// CFC twin of T_SafeMuting_Tests: the same tests drawn as CFC diagrams, the way a TwinSAFE project is authored.
    FUNCTION_BLOCK T_SafeMuting_Tests_CFC EXTENDS T_SafeCfcTestSuite
    VAR
    // Test_OssdBlockedWithoutMutingGivesSafe
    group_1 : T_SafeGroup;
    fb_1 : T_SafeMuting(group := group_1);
    // Test_SequentialMutingKeepsOutputOn
    group_2 : T_SafeGroup;
    fb_2 : T_SafeMuting(group := group_2) := (Parameters := (SequentialInputs := TRUE));
    // Test_SequenceViolationGivesError
    group_3 : T_SafeGroup;
    fb_3 : T_SafeMuting(group := group_3) := (Parameters := (SequentialInputs := TRUE));
    // Test_TwoSensorParallelSequence
    group_4 : T_SafeGroup;
    fb_4 : T_SafeMuting(group := group_4);
END_VAR

Test_OssdBlockedWithoutMutingGivesSafe();
Test_SequentialMutingKeepsOutputOn();
Test_SequenceViolationGivesError();
Test_TwoSensorParallelSequence();

METHOD PRIVATE Test_OssdBlockedWithoutMutingGivesSafe
// note: this text did not pass the execution check against the stored diagram
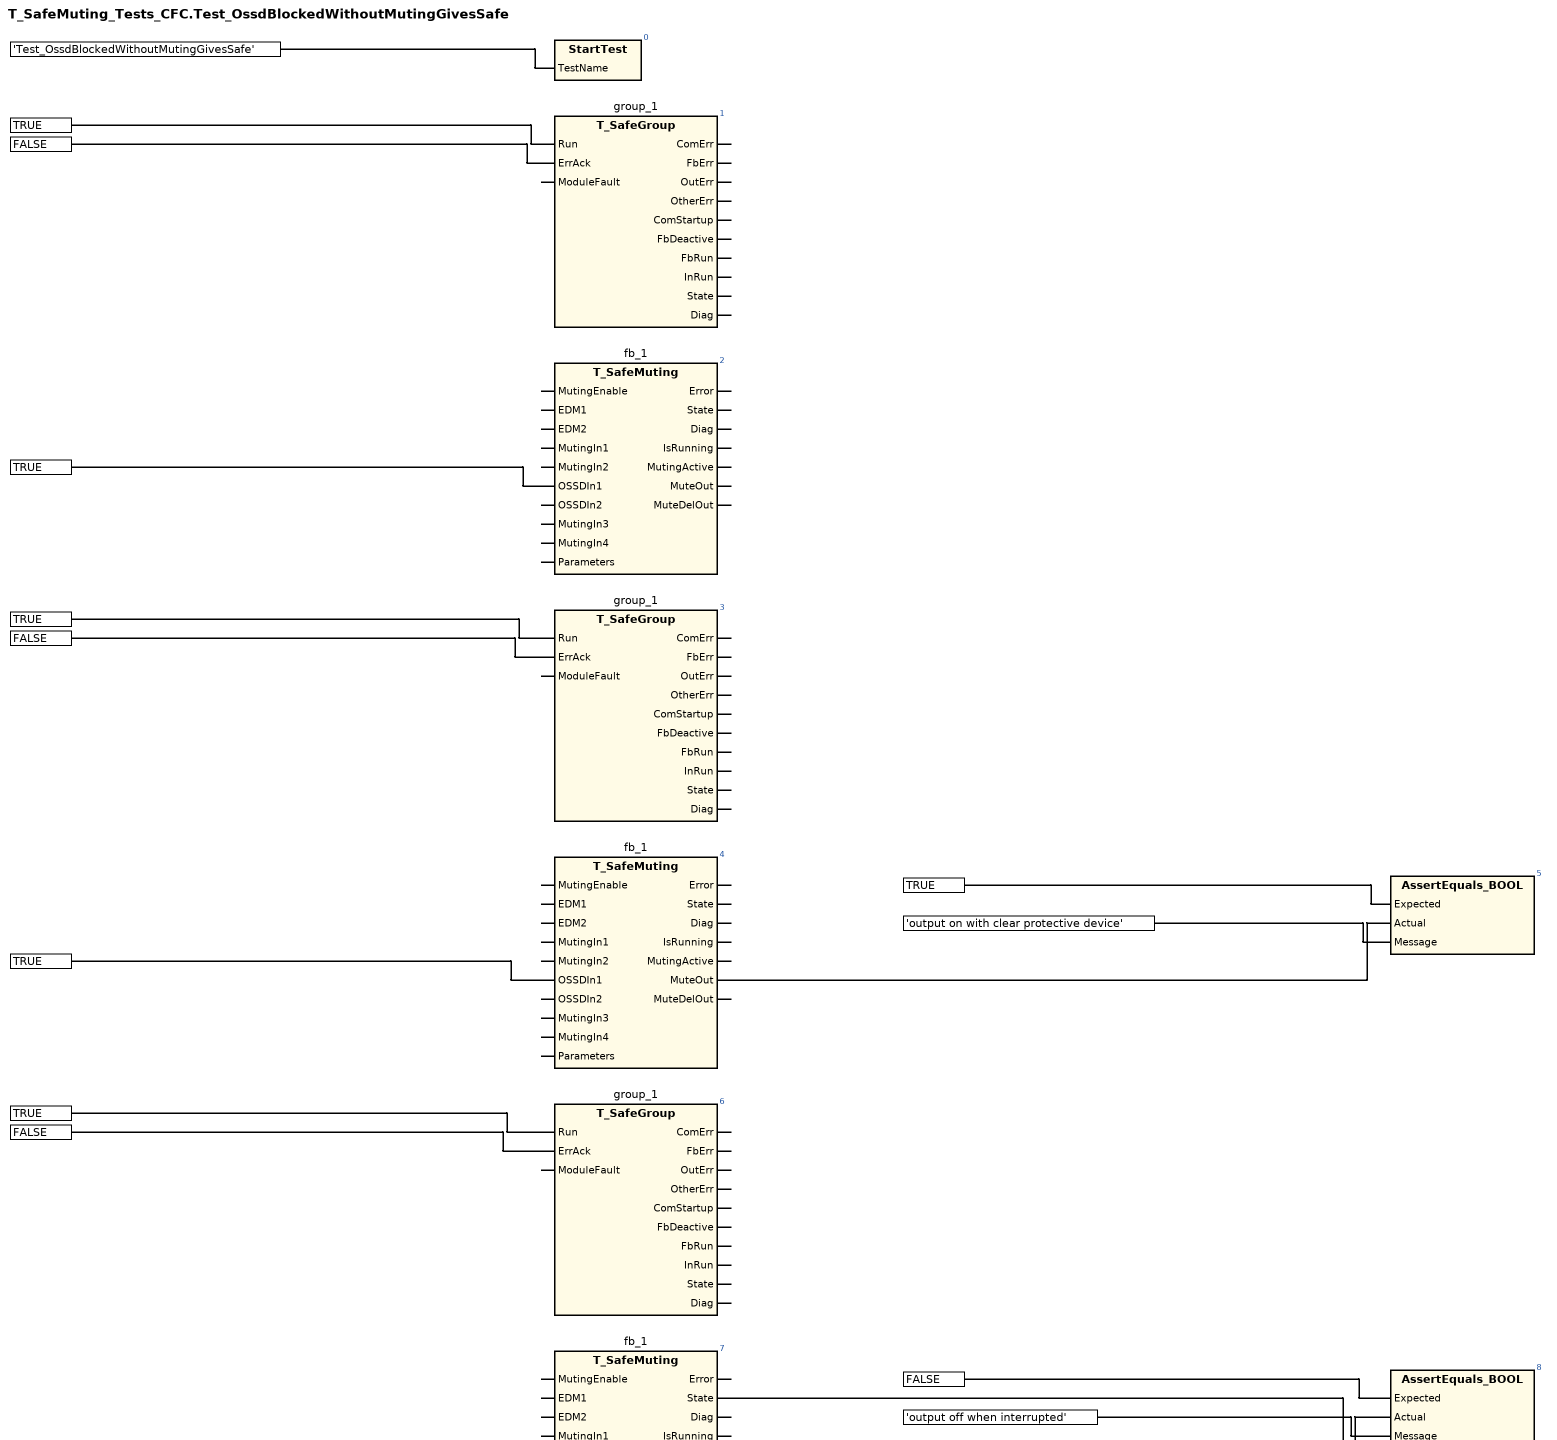
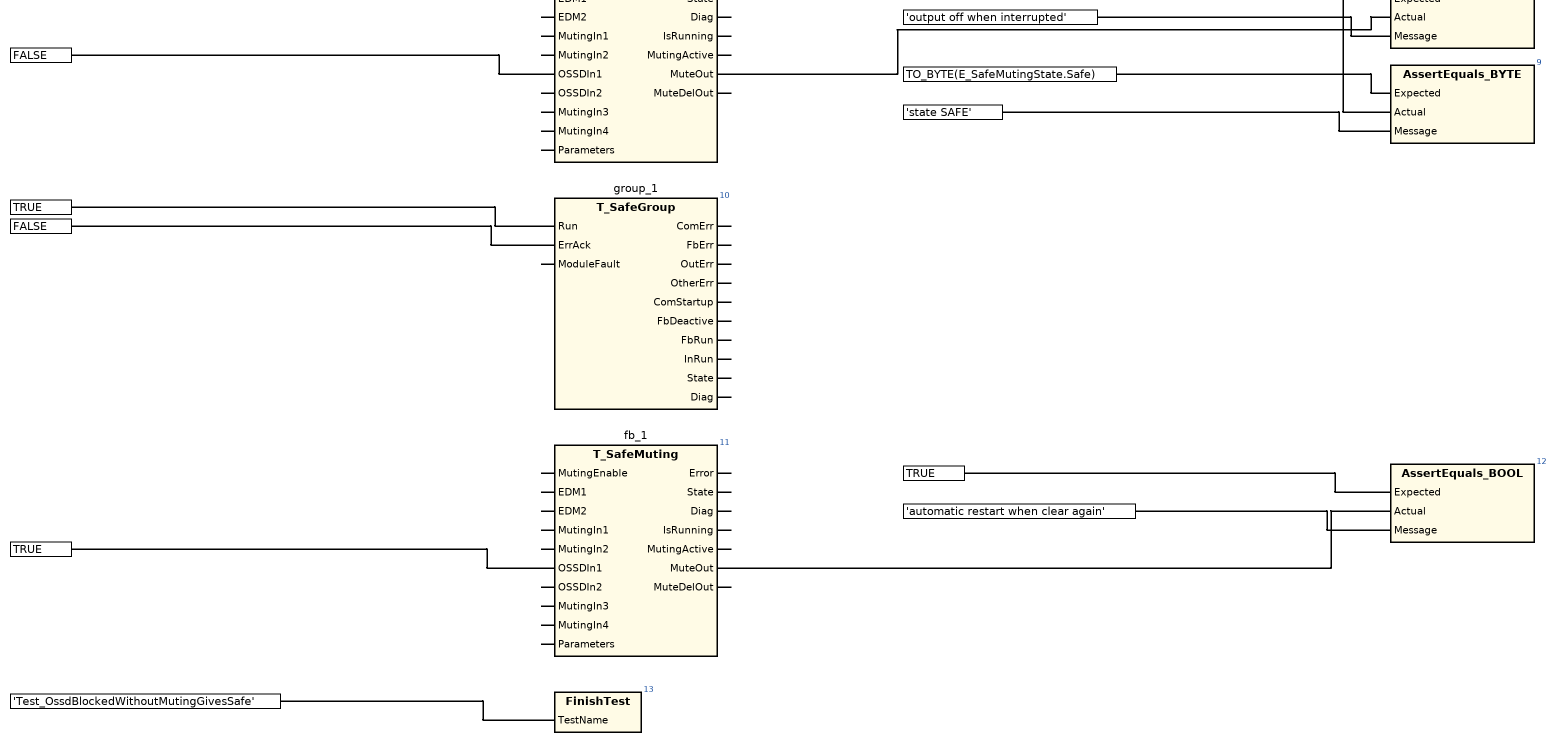
StartTest(TestName := 'Test_OssdBlockedWithoutMutingGivesSafe');
group_1(Run := TRUE, ErrAck := FALSE); // T_SafeGroup
fb_1(OSSDIn1 := TRUE); // T_SafeMuting
group_1(Run := TRUE, ErrAck := FALSE); // T_SafeGroup
fb_1(OSSDIn1 := TRUE); // T_SafeMuting
AssertEquals_BOOL(Expected := TRUE, Actual := fb_1.MuteOut, Message := 'output on with clear protective device');
group_1(Run := TRUE, ErrAck := FALSE); // T_SafeGroup
fb_1(OSSDIn1 := FALSE); // T_SafeMuting
AssertEquals_BOOL(Expected := FALSE, Actual := fb_1.MuteOut, Message := 'output off when interrupted');
AssertEquals_BYTE(Expected := TO_BYTE(E_SafeMutingState.Safe), Actual := fb_1.State, Message := 'state SAFE');
group_1(Run := TRUE, ErrAck := FALSE); // T_SafeGroup
fb_1(OSSDIn1 := TRUE); // T_SafeMuting
AssertEquals_BOOL(Expected := TRUE, Actual := fb_1.MuteOut, Message := 'automatic restart when clear again');
FinishTest(TestName := 'Test_OssdBlockedWithoutMutingGivesSafe');
END_METHOD

METHOD PRIVATE Test_SequentialMutingKeepsOutputOn
// note: this text did not pass the execution check against the stored diagram
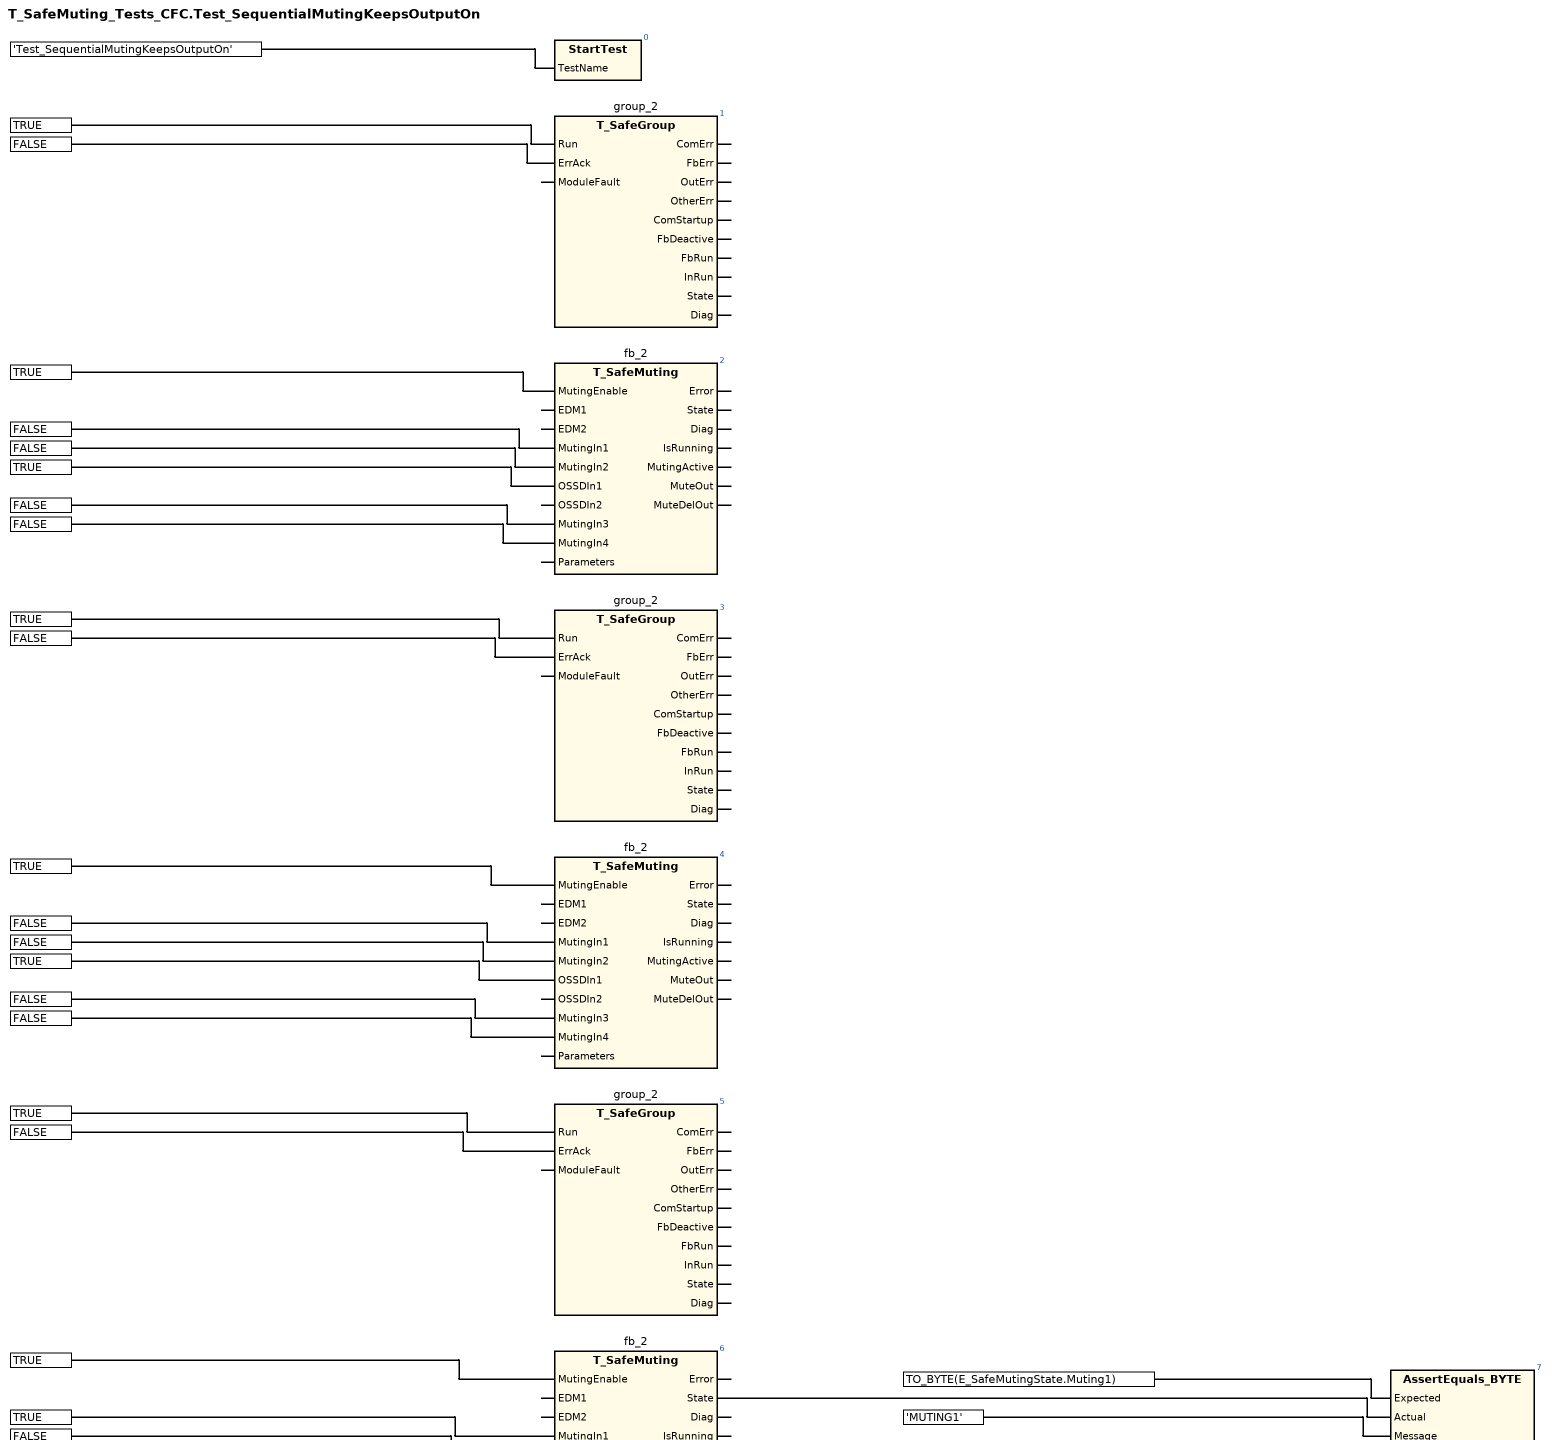
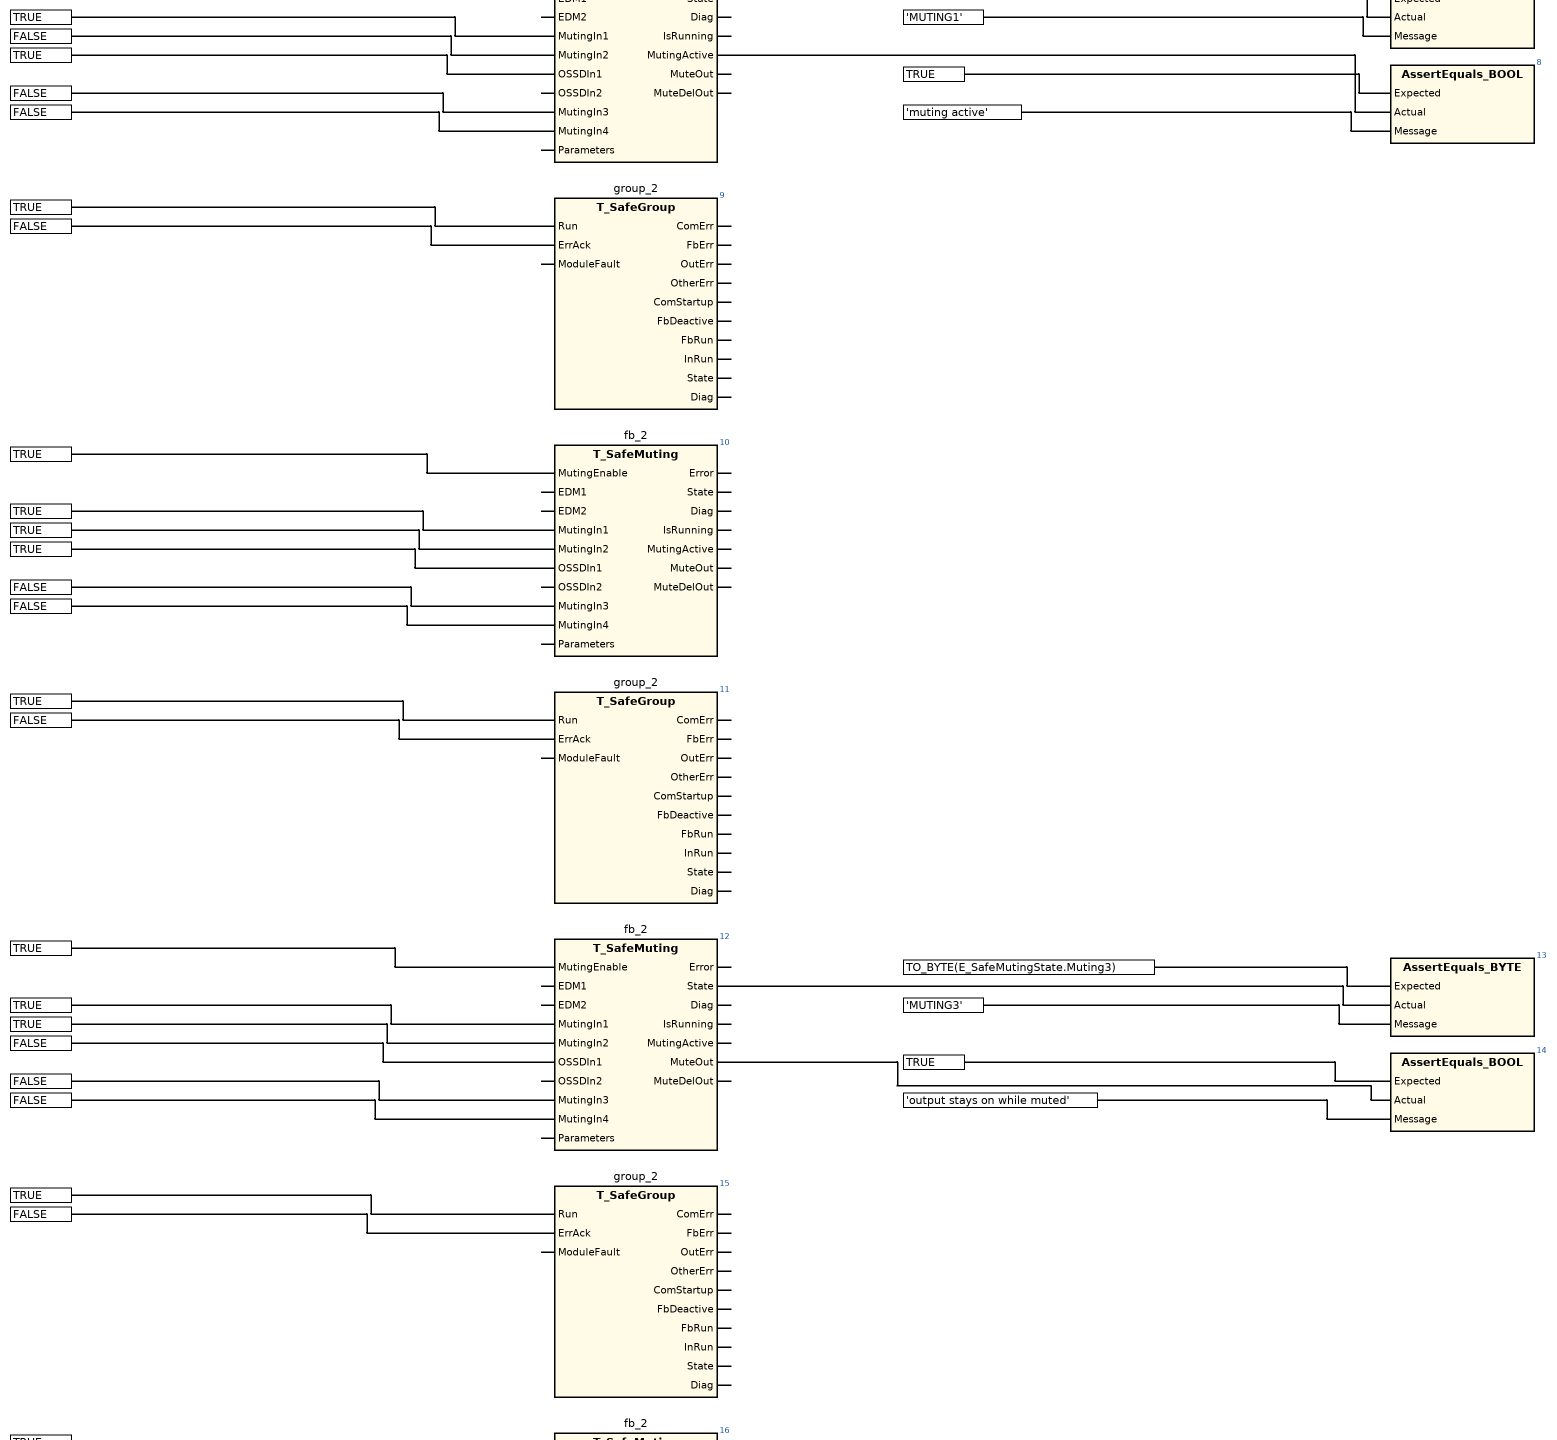
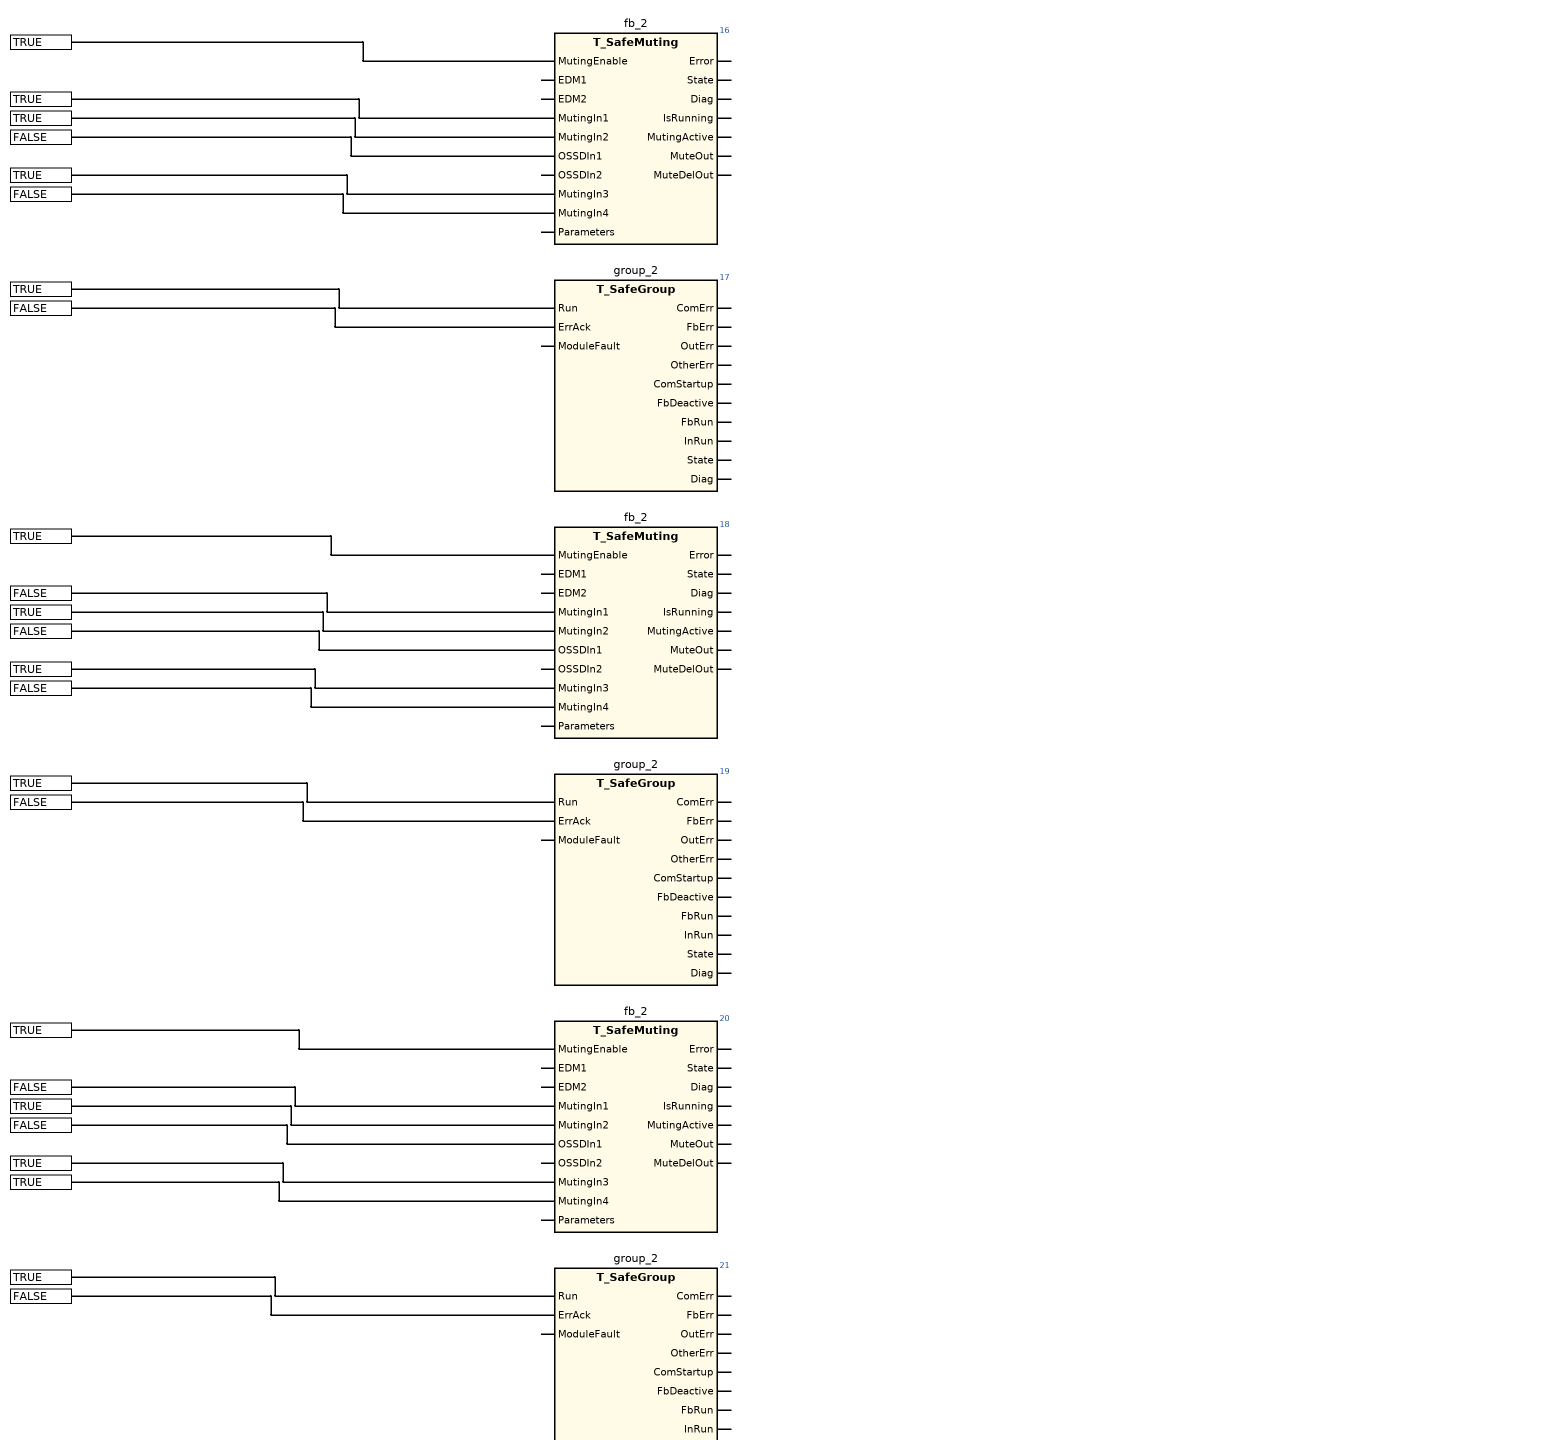
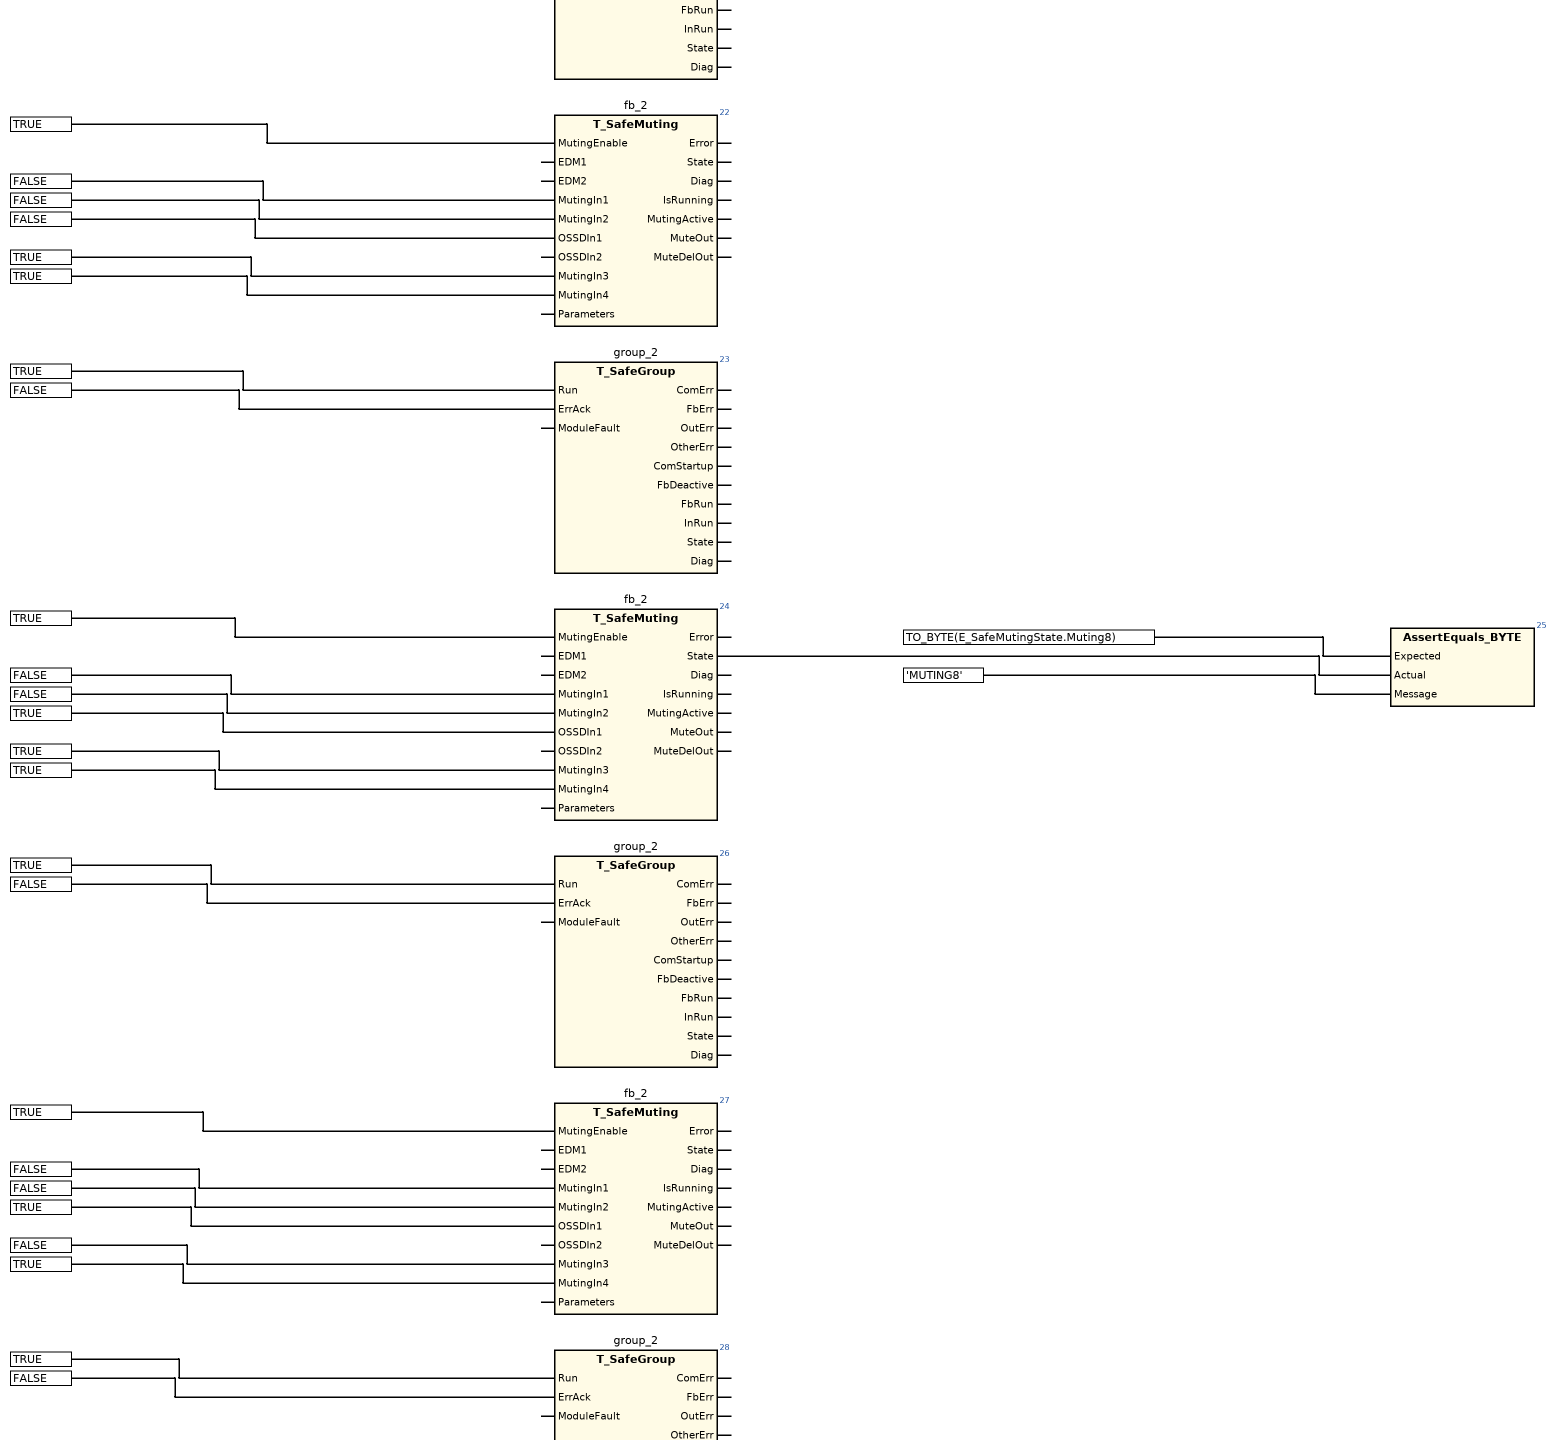
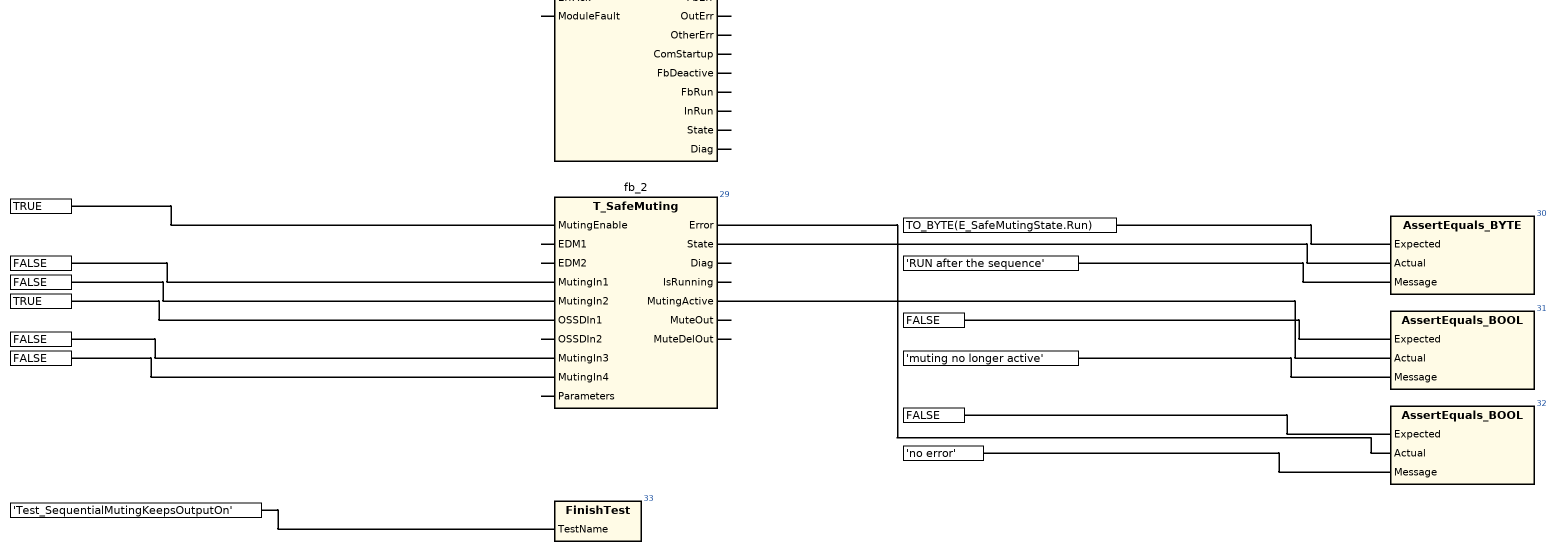
StartTest(TestName := 'Test_SequentialMutingKeepsOutputOn');
group_2(Run := TRUE, ErrAck := FALSE); // T_SafeGroup
fb_2(
    MutingEnable := TRUE,
    MutingIn1 := FALSE,
    MutingIn2 := FALSE,
    OSSDIn1 := TRUE,
    MutingIn3 := FALSE,
    MutingIn4 := FALSE); // T_SafeMuting
group_2(Run := TRUE, ErrAck := FALSE); // T_SafeGroup
fb_2(
    MutingEnable := TRUE,
    MutingIn1 := FALSE,
    MutingIn2 := FALSE,
    OSSDIn1 := TRUE,
    MutingIn3 := FALSE,
    MutingIn4 := FALSE); // T_SafeMuting
group_2(Run := TRUE, ErrAck := FALSE); // T_SafeGroup
fb_2(
    MutingEnable := TRUE,
    MutingIn1 := TRUE,
    MutingIn2 := FALSE,
    OSSDIn1 := TRUE,
    MutingIn3 := FALSE,
    MutingIn4 := FALSE); // T_SafeMuting
AssertEquals_BYTE(Expected := TO_BYTE(E_SafeMutingState.Muting1), Actual := fb_2.State, Message := 'MUTING1');
AssertEquals_BOOL(Expected := TRUE, Actual := fb_2.MutingActive, Message := 'muting active');
group_2(Run := TRUE, ErrAck := FALSE); // T_SafeGroup
fb_2(
    MutingEnable := TRUE,
    MutingIn1 := TRUE,
    MutingIn2 := TRUE,
    OSSDIn1 := TRUE,
    MutingIn3 := FALSE,
    MutingIn4 := FALSE); // T_SafeMuting
group_2(Run := TRUE, ErrAck := FALSE); // T_SafeGroup
fb_2(
    MutingEnable := TRUE,
    MutingIn1 := TRUE,
    MutingIn2 := TRUE,
    OSSDIn1 := FALSE,
    MutingIn3 := FALSE,
    MutingIn4 := FALSE); // T_SafeMuting
AssertEquals_BYTE(Expected := TO_BYTE(E_SafeMutingState.Muting3), Actual := fb_2.State, Message := 'MUTING3');
AssertEquals_BOOL(Expected := TRUE, Actual := fb_2.MuteOut, Message := 'output stays on while muted');
group_2(Run := TRUE, ErrAck := FALSE); // T_SafeGroup
fb_2(
    MutingEnable := TRUE,
    MutingIn1 := TRUE,
    MutingIn2 := TRUE,
    OSSDIn1 := FALSE,
    MutingIn3 := TRUE,
    MutingIn4 := FALSE); // T_SafeMuting
group_2(Run := TRUE, ErrAck := FALSE); // T_SafeGroup
fb_2(
    MutingEnable := TRUE,
    MutingIn1 := FALSE,
    MutingIn2 := TRUE,
    OSSDIn1 := FALSE,
    MutingIn3 := TRUE,
    MutingIn4 := FALSE); // T_SafeMuting
group_2(Run := TRUE, ErrAck := FALSE); // T_SafeGroup
fb_2(
    MutingEnable := TRUE,
    MutingIn1 := FALSE,
    MutingIn2 := TRUE,
    OSSDIn1 := FALSE,
    MutingIn3 := TRUE,
    MutingIn4 := TRUE); // T_SafeMuting
group_2(Run := TRUE, ErrAck := FALSE); // T_SafeGroup
fb_2(
    MutingEnable := TRUE,
    MutingIn1 := FALSE,
    MutingIn2 := FALSE,
    OSSDIn1 := FALSE,
    MutingIn3 := TRUE,
    MutingIn4 := TRUE); // T_SafeMuting
group_2(Run := TRUE, ErrAck := FALSE); // T_SafeGroup
fb_2(
    MutingEnable := TRUE,
    MutingIn1 := FALSE,
    MutingIn2 := FALSE,
    OSSDIn1 := TRUE,
    MutingIn3 := TRUE,
    MutingIn4 := TRUE); // T_SafeMuting
AssertEquals_BYTE(Expected := TO_BYTE(E_SafeMutingState.Muting8), Actual := fb_2.State, Message := 'MUTING8');
group_2(Run := TRUE, ErrAck := FALSE); // T_SafeGroup
fb_2(
    MutingEnable := TRUE,
    MutingIn1 := FALSE,
    MutingIn2 := FALSE,
    OSSDIn1 := TRUE,
    MutingIn3 := FALSE,
    MutingIn4 := TRUE); // T_SafeMuting
group_2(Run := TRUE, ErrAck := FALSE); // T_SafeGroup
fb_2(
    MutingEnable := TRUE,
    MutingIn1 := FALSE,
    MutingIn2 := FALSE,
    OSSDIn1 := TRUE,
    MutingIn3 := FALSE,
    MutingIn4 := FALSE); // T_SafeMuting
AssertEquals_BYTE(Expected := TO_BYTE(E_SafeMutingState.Run), Actual := fb_2.State, Message := 'RUN after the sequence');
AssertEquals_BOOL(Expected := FALSE, Actual := fb_2.MutingActive, Message := 'muting no longer active');
AssertEquals_BOOL(Expected := FALSE, Actual := fb_2.Error, Message := 'no error');
FinishTest(TestName := 'Test_SequentialMutingKeepsOutputOn');
END_METHOD

METHOD PRIVATE Test_SequenceViolationGivesError
// note: this text did not pass the execution check against the stored diagram
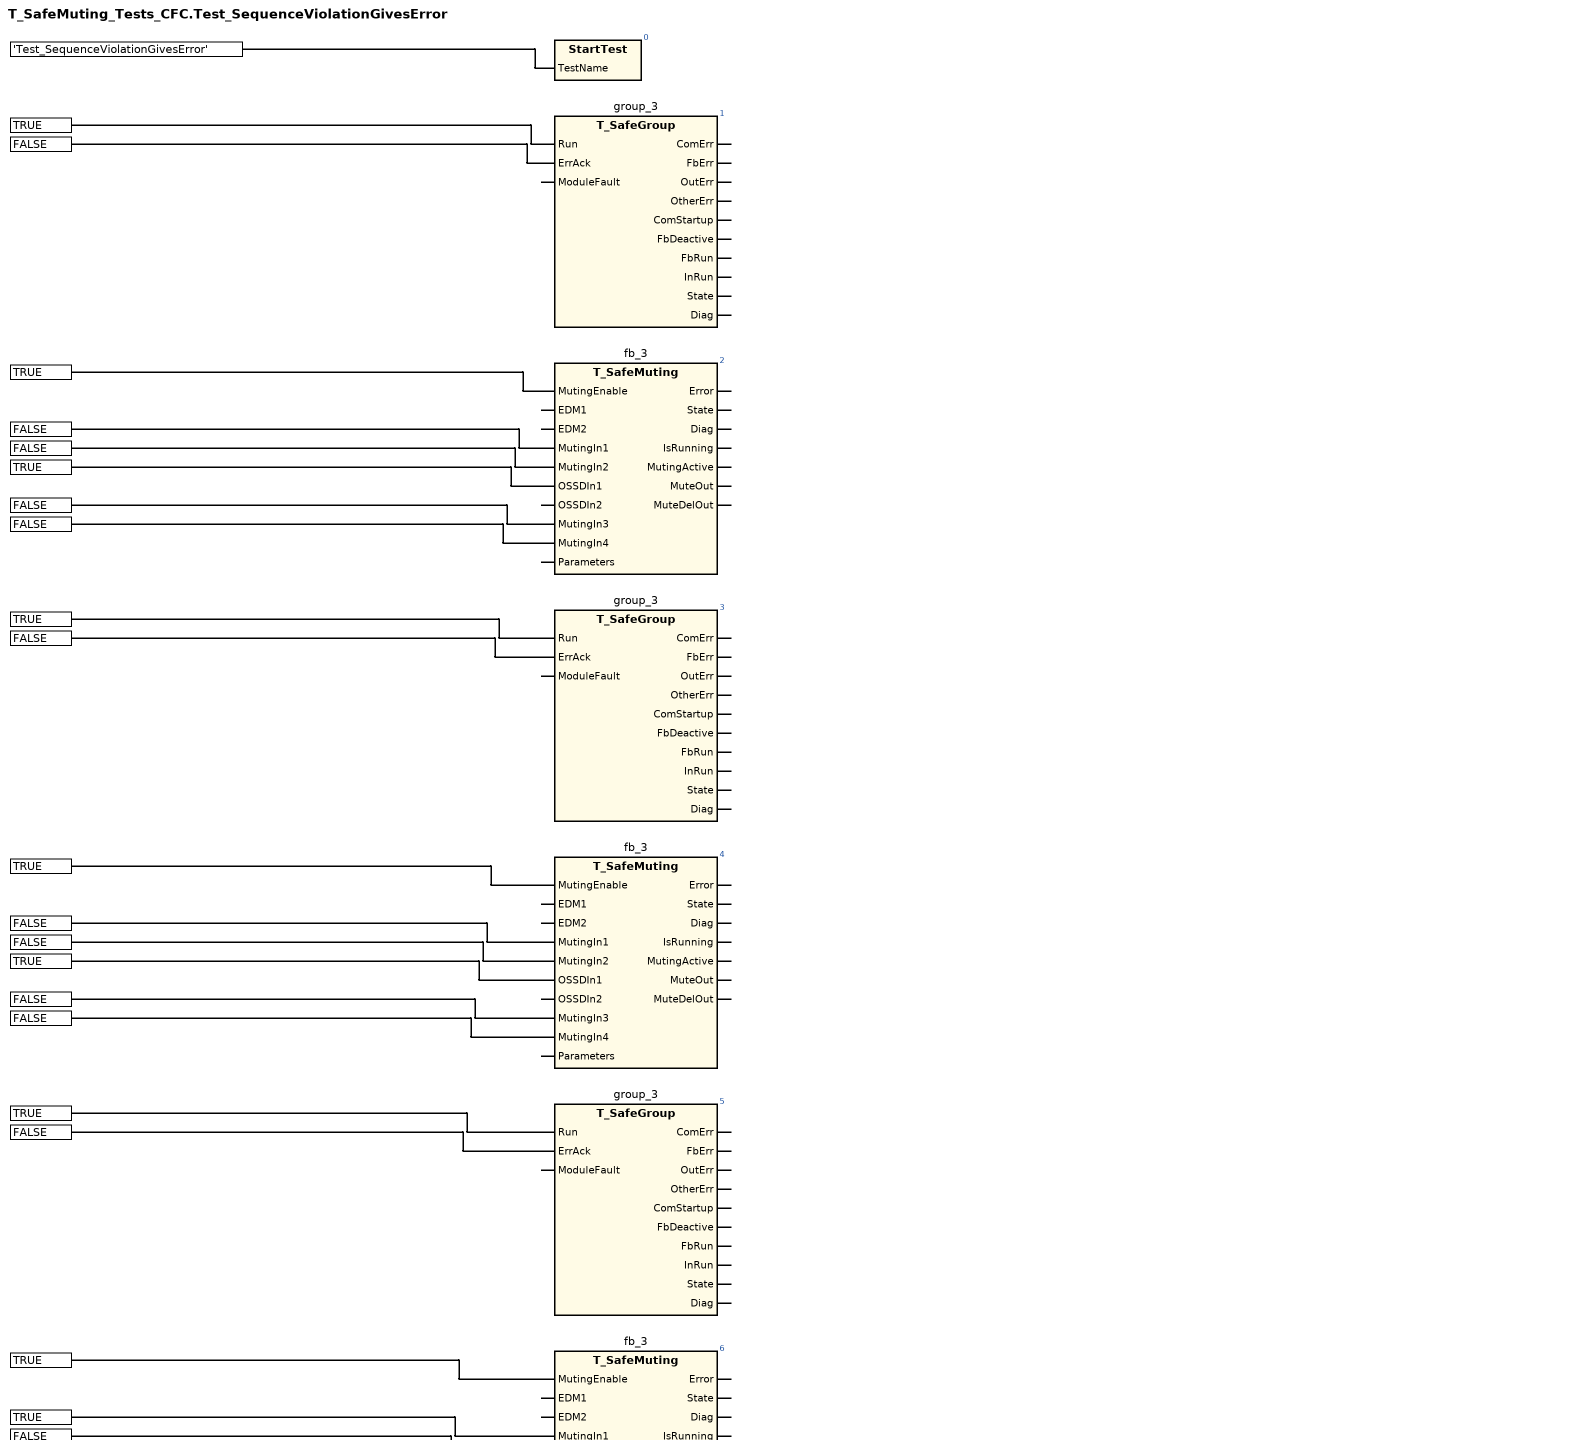
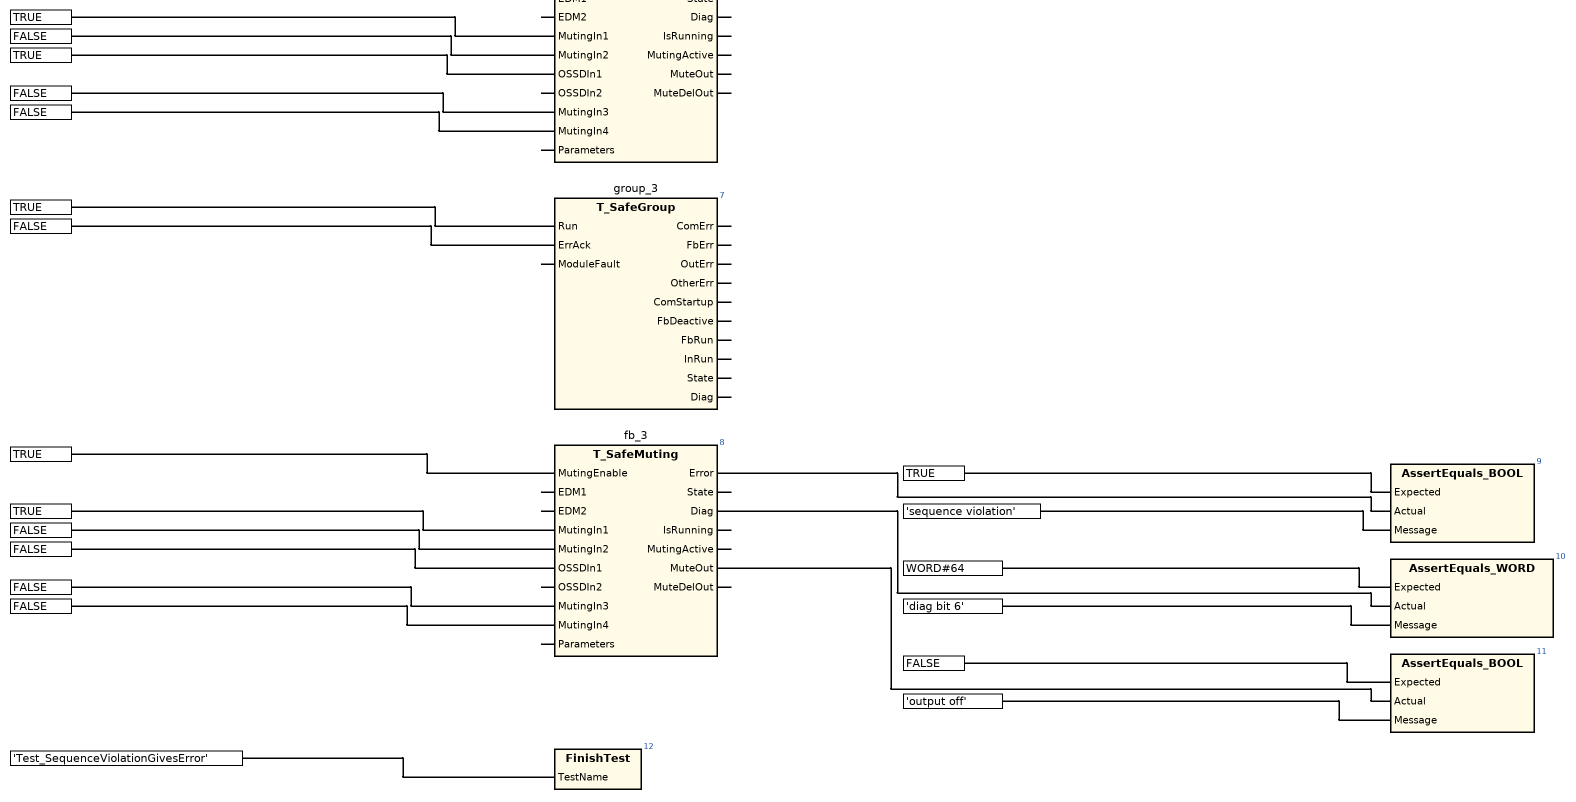
StartTest(TestName := 'Test_SequenceViolationGivesError');
group_3(Run := TRUE, ErrAck := FALSE); // T_SafeGroup
fb_3(
    MutingEnable := TRUE,
    MutingIn1 := FALSE,
    MutingIn2 := FALSE,
    OSSDIn1 := TRUE,
    MutingIn3 := FALSE,
    MutingIn4 := FALSE); // T_SafeMuting
group_3(Run := TRUE, ErrAck := FALSE); // T_SafeGroup
fb_3(
    MutingEnable := TRUE,
    MutingIn1 := FALSE,
    MutingIn2 := FALSE,
    OSSDIn1 := TRUE,
    MutingIn3 := FALSE,
    MutingIn4 := FALSE); // T_SafeMuting
group_3(Run := TRUE, ErrAck := FALSE); // T_SafeGroup
fb_3(
    MutingEnable := TRUE,
    MutingIn1 := TRUE,
    MutingIn2 := FALSE,
    OSSDIn1 := TRUE,
    MutingIn3 := FALSE,
    MutingIn4 := FALSE); // T_SafeMuting
group_3(Run := TRUE, ErrAck := FALSE); // T_SafeGroup
fb_3(
    MutingEnable := TRUE,
    MutingIn1 := TRUE,
    MutingIn2 := FALSE,
    OSSDIn1 := FALSE,
    MutingIn3 := FALSE,
    MutingIn4 := FALSE); // T_SafeMuting
AssertEquals_BOOL(Expected := TRUE, Actual := fb_3.Error, Message := 'sequence violation');
AssertEquals_WORD(Expected := WORD#64, Actual := fb_3.Diag, Message := 'diag bit 6');
AssertEquals_BOOL(Expected := FALSE, Actual := fb_3.MuteOut, Message := 'output off');
FinishTest(TestName := 'Test_SequenceViolationGivesError');
END_METHOD

METHOD PRIVATE Test_TwoSensorParallelSequence
// note: this text did not pass the execution check against the stored diagram
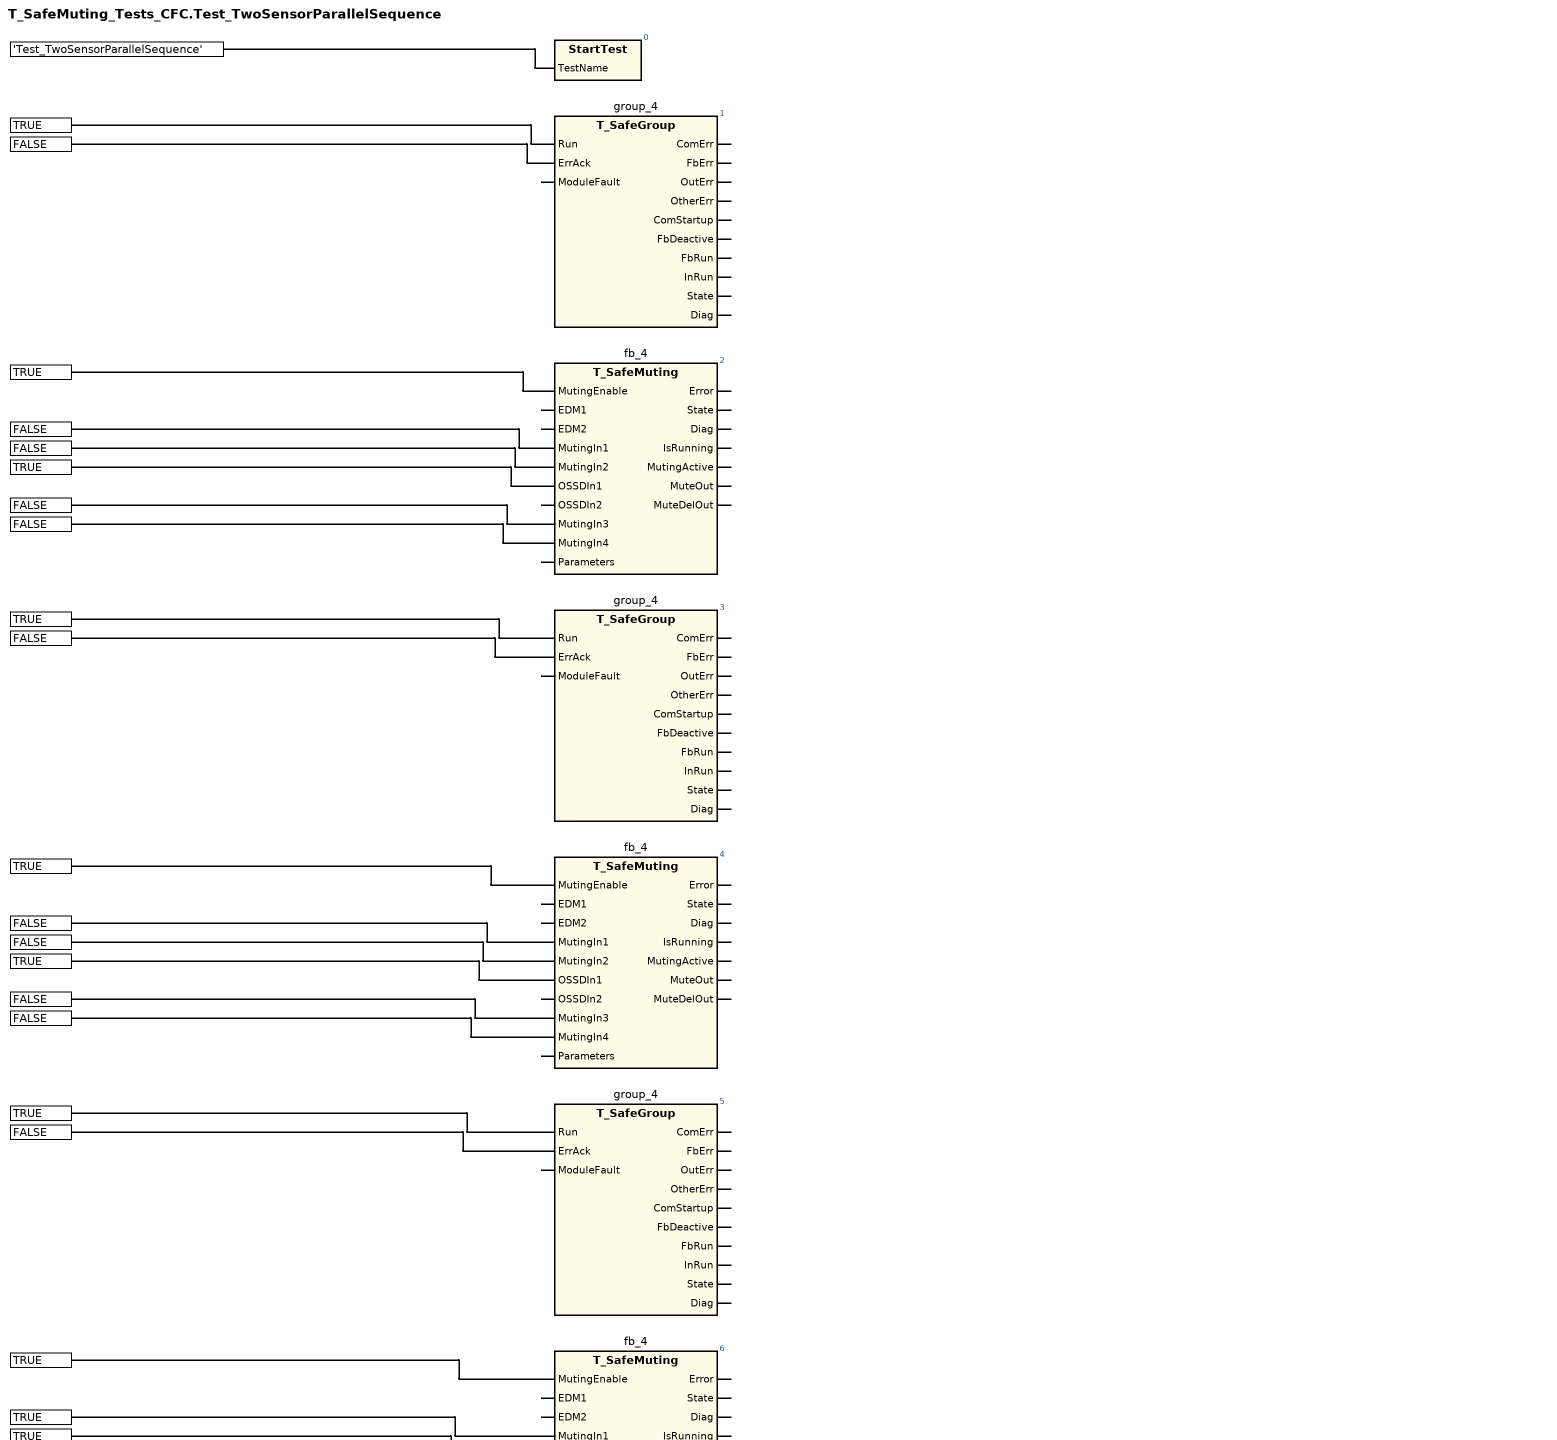
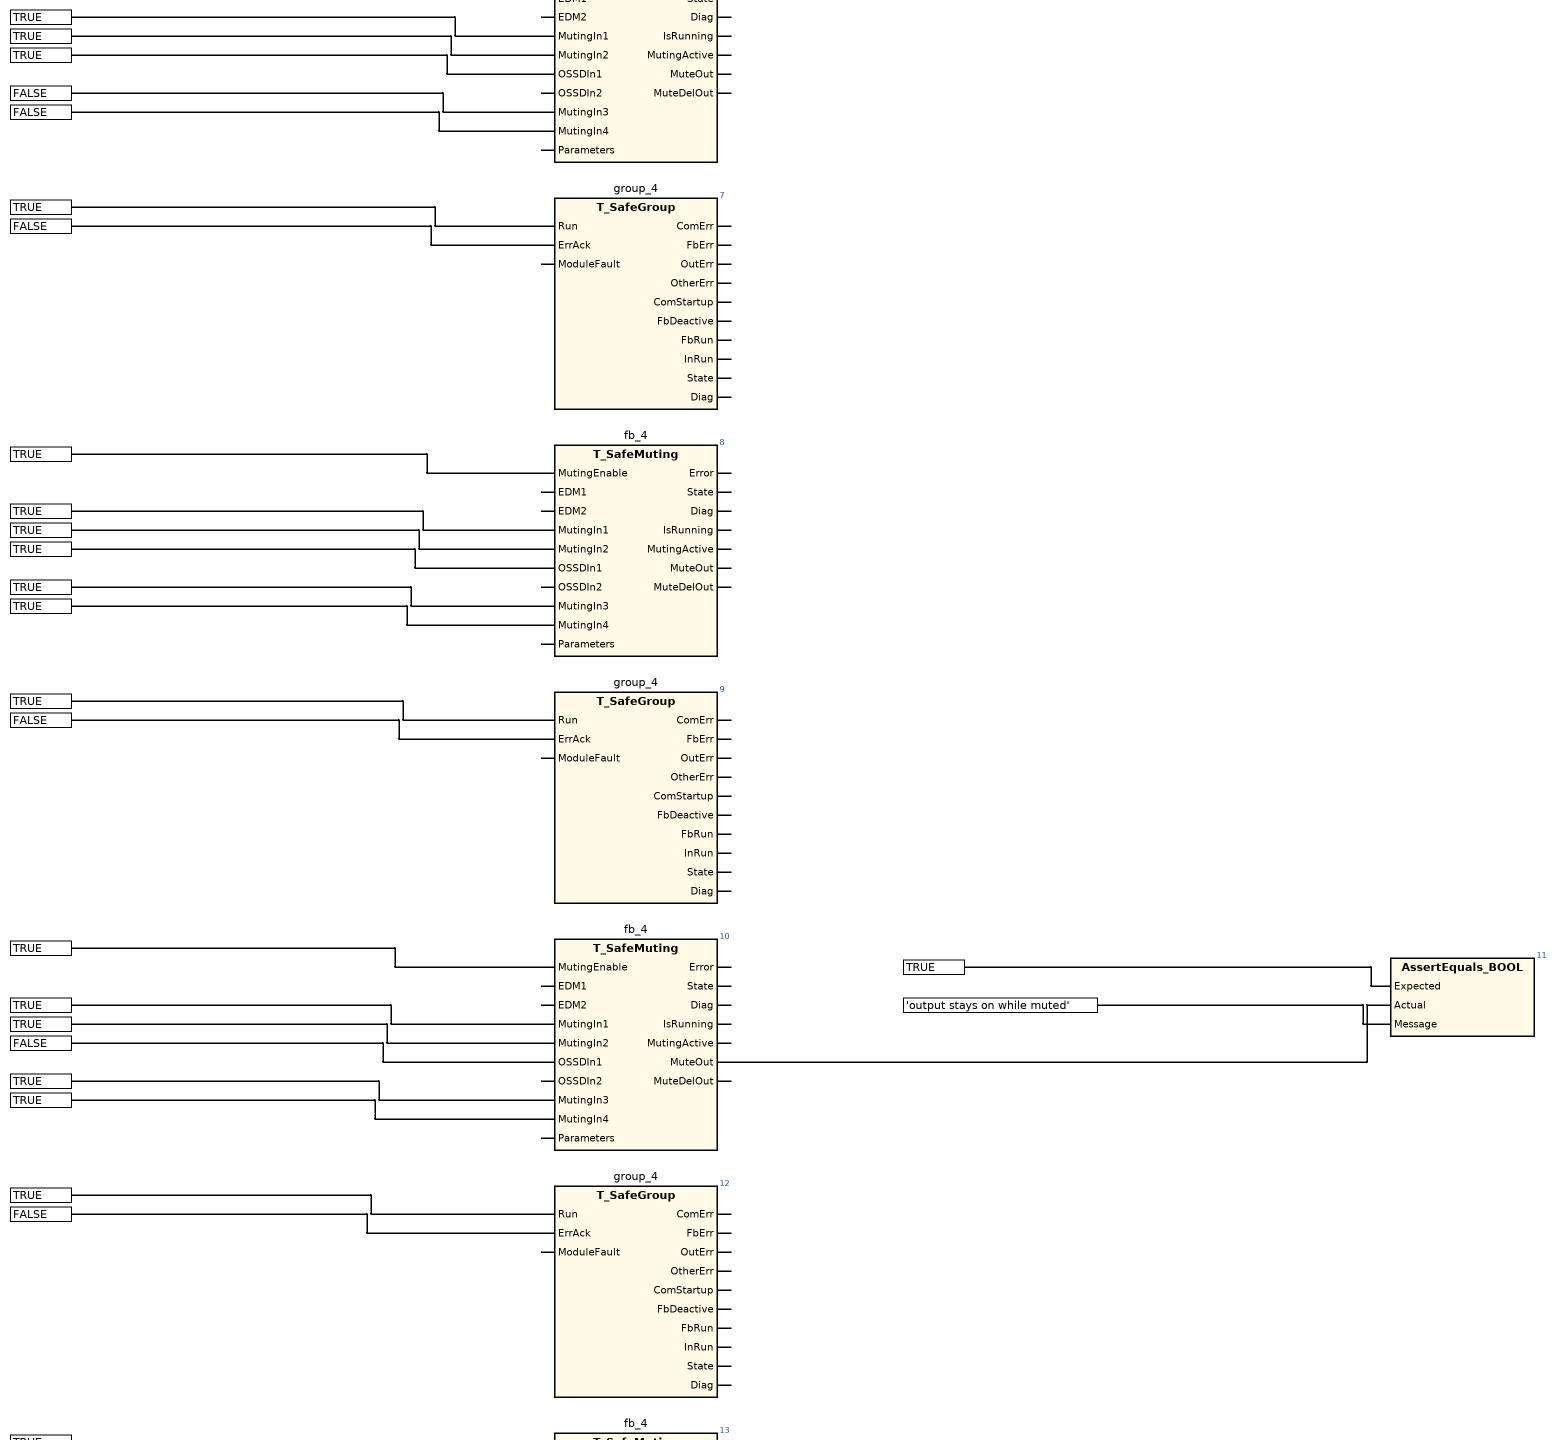
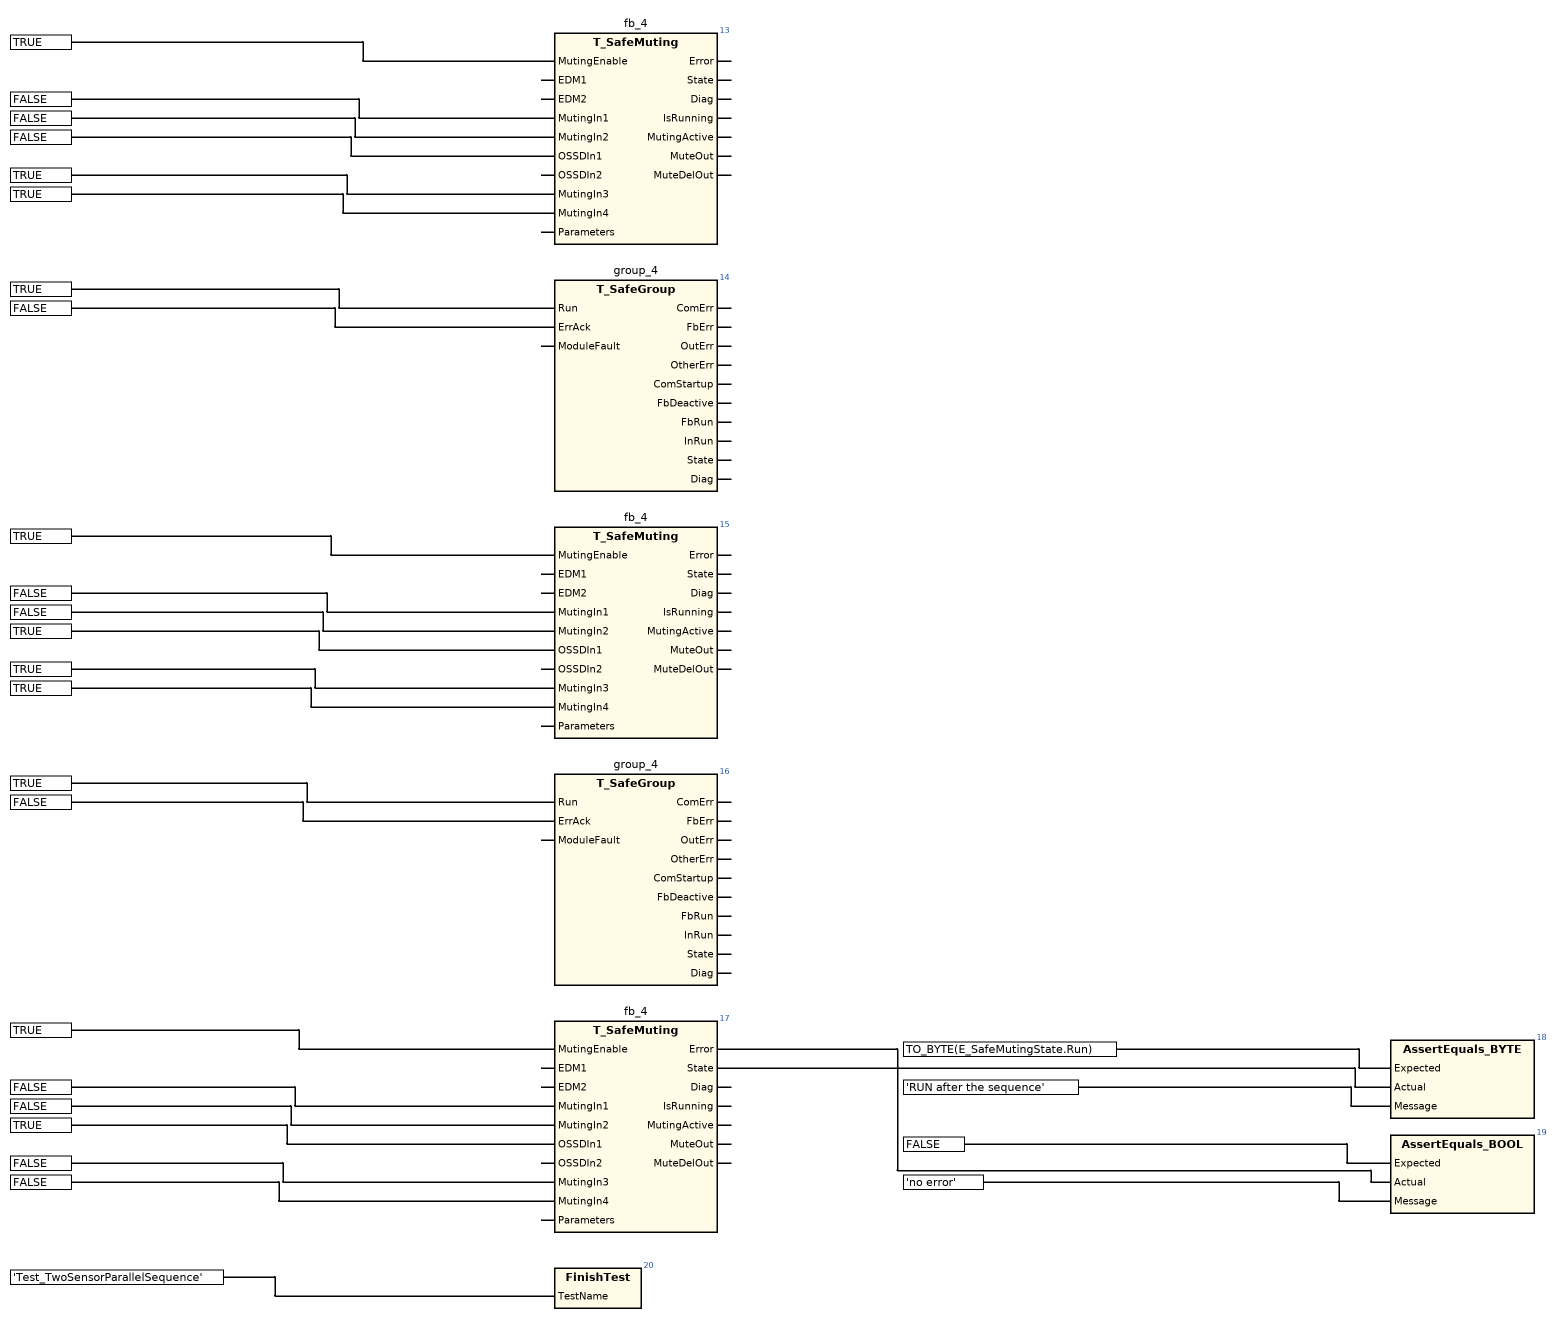
StartTest(TestName := 'Test_TwoSensorParallelSequence');
group_4(Run := TRUE, ErrAck := FALSE); // T_SafeGroup
fb_4(
    MutingEnable := TRUE,
    MutingIn1 := FALSE,
    MutingIn2 := FALSE,
    OSSDIn1 := TRUE,
    MutingIn3 := FALSE,
    MutingIn4 := FALSE); // T_SafeMuting
group_4(Run := TRUE, ErrAck := FALSE); // T_SafeGroup
fb_4(
    MutingEnable := TRUE,
    MutingIn1 := FALSE,
    MutingIn2 := FALSE,
    OSSDIn1 := TRUE,
    MutingIn3 := FALSE,
    MutingIn4 := FALSE); // T_SafeMuting
group_4(Run := TRUE, ErrAck := FALSE); // T_SafeGroup
fb_4(
    MutingEnable := TRUE,
    MutingIn1 := TRUE,
    MutingIn2 := TRUE,
    OSSDIn1 := TRUE,
    MutingIn3 := FALSE,
    MutingIn4 := FALSE); // T_SafeMuting
group_4(Run := TRUE, ErrAck := FALSE); // T_SafeGroup
fb_4(
    MutingEnable := TRUE,
    MutingIn1 := TRUE,
    MutingIn2 := TRUE,
    OSSDIn1 := TRUE,
    MutingIn3 := TRUE,
    MutingIn4 := TRUE); // T_SafeMuting
group_4(Run := TRUE, ErrAck := FALSE); // T_SafeGroup
fb_4(
    MutingEnable := TRUE,
    MutingIn1 := TRUE,
    MutingIn2 := TRUE,
    OSSDIn1 := FALSE,
    MutingIn3 := TRUE,
    MutingIn4 := TRUE); // T_SafeMuting
AssertEquals_BOOL(Expected := TRUE, Actual := fb_4.MuteOut, Message := 'output stays on while muted');
group_4(Run := TRUE, ErrAck := FALSE); // T_SafeGroup
fb_4(
    MutingEnable := TRUE,
    MutingIn1 := FALSE,
    MutingIn2 := FALSE,
    OSSDIn1 := FALSE,
    MutingIn3 := TRUE,
    MutingIn4 := TRUE); // T_SafeMuting
group_4(Run := TRUE, ErrAck := FALSE); // T_SafeGroup
fb_4(
    MutingEnable := TRUE,
    MutingIn1 := FALSE,
    MutingIn2 := FALSE,
    OSSDIn1 := TRUE,
    MutingIn3 := TRUE,
    MutingIn4 := TRUE); // T_SafeMuting
group_4(Run := TRUE, ErrAck := FALSE); // T_SafeGroup
fb_4(
    MutingEnable := TRUE,
    MutingIn1 := FALSE,
    MutingIn2 := FALSE,
    OSSDIn1 := TRUE,
    MutingIn3 := FALSE,
    MutingIn4 := FALSE); // T_SafeMuting
AssertEquals_BYTE(Expected := TO_BYTE(E_SafeMutingState.Run), Actual := fb_4.State, Message := 'RUN after the sequence');
AssertEquals_BOOL(Expected := FALSE, Actual := fb_4.Error, Message := 'no error');
FinishTest(TestName := 'Test_TwoSensorParallelSequence');
END_METHOD

END_FUNCTION_BLOCK

(* stored: Version 1.1.0.1, ProductVersion 3.1.4026.22
   POU T_SafeMuting_Tests_CFC: Id {cca67b61-3b3d-5c59-a961-95841c723a9f}, SpecialFunc None
   Method Test_OssdBlockedWithoutMutingGivesSafe: Id {a1fa14cd-f9fa-51c9-9fc1-2e15fa66dec7}
   Method Test_SequentialMutingKeepsOutputOn: Id {7fb18f84-25bf-54e2-9d32-505e87cfd692}
   Method Test_SequenceViolationGivesError: Id {45ae5d35-3403-5055-a98e-49ea11b174e7}
   Method Test_TwoSensorParallelSequence: Id {f323d194-4074-5acd-a8b1-d85ccfd714be} *)
